Staubli VAL3: getTrajList.pgx

public program getTrajList(string& x_sList[])
  local string l_sKey
begin
  resize(x_sList,1,1)
  l_sKey=first(trajTemp:tTrajItem)

  while l_sKey!=""
    x_sList[size(x_sList)-1]=l_sKey

    l_sKey=next(trajTemp:tTrajItem[l_sKey])

    if l_sKey!=""
      insert(x_sList[size(x_sList)])
    endIf
  endWhile
  if size(trajTemp:tTrajItem)<1
    x_sList=""
  endIf
end
